(* IEC 61131-3 sources: RootPLC/conformance/cases/variables, 18 files *)

(* ---- err_duplicate_pou.st ---- *)
(* spec: [variables.unique]
   expect: error RP0204 *)
TYPE Motor : STRUCT running : BOOL; END_STRUCT; END_TYPE

FUNCTION_BLOCK MOTOR
VAR_INPUT
    start : BOOL;
END_VAR
END_FUNCTION_BLOCK

(* ---- err_init_arguments_no_fb_init.st ---- *)
(* spec: [variables.init-arguments]
   expect: error RP0203 RP0119 *)
FUNCTION_BLOCK FB_Buffer
VAR_INPUT
    size : INT;
END_VAR
END_FUNCTION_BLOCK

PROGRAM PRG_Main
VAR
    b : FB_Buffer(size := 10);
END_VAR
END_PROGRAM

(* ---- err_member_named_like_variable.st ---- *)
(* spec: [variables.unique]
   expect: error RP0204 *)
FUNCTION_BLOCK Controller
VAR
    run : BOOL;
END_VAR
METHOD Run
run := TRUE;
END_METHOD
END_FUNCTION_BLOCK

(* ---- ok_init_from_local_constant.st ---- *)
(* spec: [variables.initializer] [variables.constant-names]
   expect: ok
   run: PRG_Main cycles=1
   assert: first = -1
   assert: second = -2
   assert: last = 3 *)
FUNCTION_BLOCK FB_List
VAR_OUTPUT
    current : INT := EMPTY;
    twice : INT := DOUBLE;
    top : DINT := UPPER_BOUND(items, 1);
END_VAR
VAR
    items : ARRAY[0..LAST] OF INT;
END_VAR
VAR CONSTANT
    EMPTY : INT := -1;
    DOUBLE : INT := EMPTY * 2;
    LAST : INT := 3;
END_VAR
END_FUNCTION_BLOCK

PROGRAM PRG_Main
VAR
    list : FB_List;
    first, second : INT;
    last : DINT;
END_VAR
first := list.current;
second := list.twice;
last := list.top;
END_PROGRAM

(* ---- ok_section_access.st ---- *)
(* spec: [variables.section]
   expect: ok
   run: PRG_Main cycles=1
   assert: v = 3 *)
CLASS Counter
VAR PUBLIC RETAIN
    n : INT := 3;
END_VAR
END_CLASS

PROGRAM PRG_Main
VAR
    c : Counter;
    v : INT;
END_VAR
VAR CONSTANT PUBLIC
    k : INT := 0;
END_VAR
v := c.n + k;
END_PROGRAM

(* ---- ok_var_stat_shared.st ---- *)
(* spec: [variables.static]
   expect: ok
   run: PRG_Main cycles=2
   assert: total = 6
   assert: mine = 2 *)
FUNCTION_BLOCK FB_Shared
VAR_OUTPUT
    calls : INT;
    own : INT;
END_VAR
VAR_STAT
    shared : INT;
END_VAR
shared := shared + 1;
own := own + 1;
calls := shared;
END_FUNCTION_BLOCK

PROGRAM PRG_Main
VAR
    a, b : FB_Shared;
    total, mine : INT;
END_VAR
a();
b();
b();
total := b.calls;
mine := a.own;
END_PROGRAM

(* ---- warn_fb_initializer.st ---- *)
(* spec: [variables.initializer] [scope.vendor-forms]
   expect: warning RP0134
   run: PRG_Main cycles=1
   assert: pt = T#1S
   assert: n = 7
   assert: d = 3 *)
FUNCTION_BLOCK FB_Count
VAR_INPUT
    k : INT := 3;
END_VAR
VAR_OUTPUT
    Count : INT;
END_VAR
Count := k;
END_FUNCTION_BLOCK

PROGRAM PRG_Main
VAR
    t : TON := (PT := T#1S);
    a : FB_Count := (k := 7);
    b : FB_Count := ();
    pt : TIME;
    n, d : INT;
END_VAR
a();
b();
pt := t.PT;
n := a.Count;
d := b.Count;
END_PROGRAM

(* ---- warn_init_arguments.st ---- *)
(* spec: [variables.init-arguments] [pous.oop.fb-init]
   expect: warning RP0119 RP0135
   run: PRG_Main cycles=1
   assert: small = 10
   assert: named = 'B2'
   assert: parent_ok = TRUE *)
FUNCTION_BLOCK FB_Buffer
VAR_OUTPUT
    size : INT;
    name : STRING;
    hasParent : BOOL;
END_VAR
METHOD FB_init : BOOL
VAR_INPUT
    bInitRetains : BOOL;
    bInCopyCode : BOOL;
    nSize : INT;
    sName : STRING;
    ipParent : REF_TO PRG_Main;
END_VAR
size := nSize;
name := sName;
hasParent := ipParent <> NULL;
END_METHOD
END_FUNCTION_BLOCK

PROGRAM PRG_Main
VAR
    a : FB_Buffer(10, 'A1');
    b : FB_Buffer(sName := 'B2', nSize := 20, ipParent := REF(THIS^));
    small : INT;
    named : STRING;
    parent_ok : BOOL;
END_VAR
small := a.size;
named := b.name;
parent_ok := b.hasParent AND NOT a.hasParent;
END_PROGRAM

(* ---- warn_init_from_variable.st ---- *)
(* spec: [variables.initializer.variable] [scope.vendor-forms]
   expect: warning RP0135
   run: PRG_Main cycles=1
   assert: left = 6000
   assert: half = 3000
   assert: early = 0
   assert: fromFun = 12 *)
FUNCTION_BLOCK Tank
VAR_OUTPUT
    early : DINT := later;
    maxMs : DINT := 6000;
    leftMs : DINT := maxMs;
    halfMs : DINT := maxMs / 2;
    later : DINT := 7;
END_VAR
leftMs := leftMs;
END_FUNCTION_BLOCK

FUNCTION Twice : DINT
VAR_INPUT
    x : DINT;
END_VAR
VAR
    base : DINT := 6;
    double : DINT := base * 2;
END_VAR
Twice := double + x * 0;
END_FUNCTION

PROGRAM PRG_Main
VAR
    t : Tank;
    left, half, early, fromFun : DINT;
END_VAR
t();
left := t.leftMs;
half := t.halfMs;
early := t.early;
fromFun := Twice(1);
END_PROGRAM

(* ---- err_duplicate_name.st ---- *)
(* spec: [variables.unique]
   expect: error RP0204 *)
PROGRAM PRG_Main
VAR_INPUT
    speed : INT;
END_VAR
VAR
    SPEED : REAL;
END_VAR
END_PROGRAM

(* ---- err_initializer_type.st ---- *)
(* spec: [variables.initializer.check]
   expect: error RP0103 *)
PROGRAM PRG_Main
VAR
    b : BOOL := 'on';
END_VAR
END_PROGRAM

(* ---- err_unknown_member.st ---- *)
(* spec: [variables.resolution]
   expect: error RP0203 *)
PROGRAM PRG_Main
VAR
    tmr : TON;
    b : BOOL;
END_VAR
b := tmr.QQ;
END_PROGRAM

(* ---- err_unknown_name.st ---- *)
(* spec: [variables.resolution]
   expect: error RP0203 *)
PROGRAM PRG_Main
VAR
    x : INT;
END_VAR
x := y + 1;
END_PROGRAM

(* ---- ok_initializers.st ---- *)
(* spec: [variables.initializer]
   expect: ok
   run: PRG_Main cycles=1
   assert: a[2] = 3
   assert: p.y = 2 *)
TYPE Point : STRUCT x : INT; y : INT; END_STRUCT; END_TYPE

PROGRAM PRG_Main
VAR
    a : ARRAY[0..2] OF INT := [1, 2, 3];
    p : Point := (x := 1, y := 2);
END_VAR
END_PROGRAM

(* ---- ok_located.st ---- *)
(* spec: [variables.located]
   expect: ok *)
PROGRAM PRG_Main
VAR
    button AT %IX0.0 : BOOL;
    lamp AT %QX0.1 : BOOL;
END_VAR
lamp := button;
END_PROGRAM

(* ---- ok_resolution.st ---- *)
(* spec: [variables.resolution] [variables.initializer.check]
   expect: ok
   run: PRG_Main cycles=1
   assert: n = 5 *)
TYPE Pt : STRUCT x : INT; y : INT; END_STRUCT; END_TYPE
TYPE Color : (Red, Green); END_TYPE

FUNCTION Twice : INT
VAR_INPUT
    v : INT;
END_VAR
Twice := v * 2;
END_FUNCTION

PROGRAM PRG_Main
VAR
    p : Pt := (x := 1);
    c : Color := Green;
    k : ARRAY[1..3] OF INT := [1, 2, 3];
    n : INT;
END_VAR
n := Twice(p.x) + k[3];
END_PROGRAM

(* ---- ok_sections.st ---- *)
(* spec: [variables.section] [variables.declaration] [pous.program] [syntax.pragmas]
   expect: ok *)
PROGRAM PRG_Main
VAR_INPUT
    start, stop : BOOL;
END_VAR
VAR_OUTPUT
    running : BOOL;
END_VAR
VAR CONSTANT
    LIMIT : INT := 10;
END_VAR
VAR RETAIN
    {attribute 'hide'}
    count : DINT;
END_VAR
running := (start OR running) AND NOT stop;
END_PROGRAM

(* ---- warn_array_init_repeat.st ---- *)
(* spec: [variables.initializer] [scope.vendor-forms]
   expect: warning RP0135
   run: PRG_Main cycles=1
   assert: a[0] = 1
   assert: a[1] = 7
   assert: a[3] = 7
   assert: a[4] = 2
   assert: a[5] = 0
   assert: d[2] = 0
   assert: d[3] = 9
   assert: e[2] = 5 *)
PROGRAM PRG_Main
VAR
    a : ARRAY[0..5] OF INT := [1, 3(7), 2];   (* 3(7): three elements of 7 *)
    d : ARRAY[0..3] OF INT := [1, 2(), 9];    (* 2(): two defaults *)
    e : ARRAY[0..2] OF INT := [(1 + 2)(5)];   (* a constant expression as count *)
END_VAR
END_PROGRAM
